(* PLC project globals, tcpethernet globals 1 *)
(* stored: creationDateTime 2026-11-15T09:00:00, modificationDateTime 2026-11-15T09:00:00 *)

FUNCTION_BLOCK Bump
  VAR_INPUT
    amount : DINT;
  END_VAR
  VAR_EXTERNAL
    ResourceGlobal : DINT;
  END_VAR

            ResourceGlobal := ResourceGlobal + amount;
          
END_FUNCTION_BLOCK

PROGRAM plc_prg
  VAR
    b : Bump;
    seen : DINT;
    limit_seen : INT;
  END_VAR
  VAR_EXTERNAL CONSTANT
    ResetCounterValue : INT;
  END_VAR

            b(amount := 3);
seen := ResourceGlobal;
limit_seen := ResetCounterValue;
Hits := Hits + 1;
          
END_PROGRAM

CONFIGURATION config
  VAR_GLOBAL CONSTANT
    ResetCounterValue : INT := 17;
  END_VAR
  VAR_GLOBAL RETAIN
    Hits : DINT;
  END_VAR
  RESOURCE resource1 ON PLC
    VAR_GLOBAL
      ResourceGlobal : DINT := 2;
    END_VAR
    TASK task0(INTERVAL := T#20ms, PRIORITY := 0);
    PROGRAM instance0 WITH task0 : plc_prg;
  END_RESOURCE
END_CONFIGURATION
